{region 'Documentation'}
(*!
<summary>Checks that the rising-edge count is less than or equal to the maximum.</summary>
<description>

Observation and accumulated-count handling come from AssertionEdgeCountBase. Evaluate
checks the held count independently of Enable; reset clears the count and baseline.

</description>
*)
{endregion}
FUNCTION_BLOCK AssertRisingEdgeCntLessEqual EXTENDS AssertionEdgeCountBase
VAR_INPUT
    Maximum : UINT; //! Inclusive upper bound of the comparison; for a range, must not be below Minimum.
END_VAR

SUPER^();

{region 'Documentation'}
(*!
<summary>Observe through the base, then evaluate the count with Error priority.</summary>
*)
{endregion}
METHOD PROTECTED Assert
VAR
    Message : STRING(GVL_Constants.MessageLength);
    MaximumText : STRING(GVL_Constants.AssertionValueLength);
    ActualText : STRING(GVL_Constants.AssertionValueLength);
END_VAR
SUPER^.Assert();

IF NOT EvaluationActive THEN
    RETURN;
END_IF;

IF Result = E_Result.Error THEN
    RETURN;
END_IF;

IF Result = E_Result.Failed THEN
    RETURN;
END_IF;

IF EdgeCount > Maximum THEN
    MaximumText := UINT_TO_STRING(Maximum);
    ActualText := UINT_TO_STRING(EdgeCount);
    Message := CONCAT('Assertion failed: rising edge count is above maximum. Maximum = ',
        MaximumText);
    Message := CONCAT(Message, ', Actual = ');
    Message := CONCAT(Message, ActualText);
    Message := CONCAT(Message, '.');
    Fail(Message := Message);
    RETURN;
END_IF;

Pass();
END_METHOD

{region 'Documentation'}
(*!
<summary>Recognize a rising edge without changing observation state.</summary>
*)
{endregion}
METHOD PROTECTED IsMatchingEdge : BOOL //! TRUE when PreviousValue and CurrentValue form the edge selected by this Assertion.
VAR_INPUT
    PreviousValue : BOOL; //! Signal value from the preceding active observation.
    CurrentValue : BOOL; //! Signal value from the current active observation.
END_VAR
IsMatchingEdge := NOT PreviousValue AND CurrentValue;
END_METHOD

END_FUNCTION_BLOCK

(* stored: Version 1.1.0.1
   POU AssertRisingEdgeCntLessEqual: Id {9b664c90-9a37-4878-befc-48e7039f8775}, SpecialFunc None
   Folder Internal: Id {cc7978f7-8929-4c93-a731-e9f09955db04}
   Method Assert: Id {21715219-e411-4e65-bf17-6d1daef5378c}
   Method IsMatchingEdge: Id {fc8c36cd-228b-40ab-9b53-9c246ac6a7c5} *)
